SUBAPPLICATION SubApp_PC_B (* Geraet B: Variablen per CLIENT (opcua.adoc): Input_I1 schreibt 42 auf Increment (CLIENT_1_0), liest danach Incremented = 43 (CLIENT_0_1) *)
  (* Standard: 61499-2; Description: Copyright (c) 2026 Meisterschulen am Ostbahnhof This program and the accompanying materials are made available under the terms of the Eclipse Public License 2.0 which is available at https://www.eclipse.org/legal/epl-2.0/ SPDX-License-Identifier: EPL-2.0 *)
  (* Version 1.0, 2026-10-18, Franz Höpfinger, Meisterschulen am Ostbahnhof, opcua.adoc-Beispiel auf zwei Geraeten *)
  PACKAGE subapp::Training_16_OPC_UA_RES;
  IMPORT VV::const::OPC_UA::myOpcUaAddresses::T16_INC_READ;
  IMPORT VV::const::OPC_UA::myOpcUaAddresses::T16_INCD_WRITE;
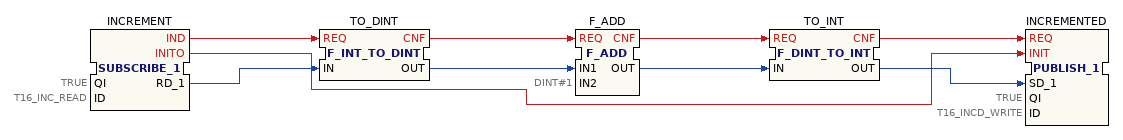
  FBS
    INCREMENT : iec61499::net::SUBSCRIBE_1(QI := TRUE, ID := T16_INC_READ);
    TO_DINT : iec61131::conversion::F_INT_TO_DINT;
    F_ADD : iec61131::arithmetic::F_ADD(IN2 := DINT#1);
    TO_INT : iec61131::conversion::F_DINT_TO_INT;
    INCREMENTED : iec61499::net::PUBLISH_1(QI := TRUE, ID := T16_INCD_WRITE);
  END_FBS
  EVENT_CONNECTIONS
    INCREMENT.IND TO TO_DINT.REQ;
    TO_DINT.CNF TO F_ADD.REQ;
    F_ADD.CNF TO TO_INT.REQ;
    TO_INT.CNF TO INCREMENTED.REQ;
    INCREMENT.INITO TO INCREMENTED.INIT;
  END_CONNECTIONS
  DATA_CONNECTIONS
    INCREMENT.RD_1 TO TO_DINT.IN;
    TO_DINT.OUT TO F_ADD.IN1;
    F_ADD.OUT TO TO_INT.IN;
    TO_INT.OUT TO INCREMENTED.SD_1;
  END_CONNECTIONS
END_SUBAPPLICATION
